TYPE "DT_ALM_SYSTEM_GEN_SPEED_WH_AND_VIB"
VERSION : 0.1
   STRUCT
      F1_ERR { S7_SetPoint := 'False'} : "DT_ALM_SOLO" := (192, FALSE, FALSE, TRUE, (), (), 2, 4, 2, (), (), (), (), (), T#3S);
      F1_H { S7_SetPoint := 'False'} : "DT_ALM_SOLO" := (193, FALSE, FALSE, TRUE, (), (), 2, 4, 1, (), (), (), (), (), T#5S);
      F1_HH { S7_SetPoint := 'False'} : "DT_ALM_SOLO" := (194, FALSE, FALSE, TRUE, (), (), 2, 4, 3, (), (), (), (), (), T#5S);
      F2_ERR { S7_SetPoint := 'False'} : "DT_ALM_SOLO" := (195, FALSE, FALSE, TRUE, (), (), 2, 4, 2, (), (), (), (), (), T#3S);
      F2_H { S7_SetPoint := 'False'} : "DT_ALM_SOLO" := (196, FALSE, FALSE, TRUE, (), (), 2, 4, 1, (), (), (), (), (), T#5S);
      F2_HH { S7_SetPoint := 'False'} : "DT_ALM_SOLO" := (197, FALSE, FALSE, TRUE, (), (), 2, 4, 3, (), (), (), (), (), T#5S);
      F3_ERR { S7_SetPoint := 'False'} : "DT_ALM_SOLO" := (198, FALSE, FALSE, FALSE, (), (), 0, 0, 0, (), (), (), (), (), T#500MS);
      F3_H { S7_SetPoint := 'False'} : "DT_ALM_SOLO" := (199, FALSE, FALSE, FALSE, (), (), 0, 0, 0, (), (), (), (), (), T#500MS);
      F3_HH { S7_SetPoint := 'False'} : "DT_ALM_SOLO" := (200, FALSE, FALSE, FALSE, (), (), 0, 0, 0, (), (), (), (), (), T#500MS);
      F4_ERR { S7_SetPoint := 'False'} : "DT_ALM_SOLO" := (201, FALSE, FALSE, TRUE, (), (), 2, 4, 2, (), (), (), (), (), T#3S);
      F4_H { S7_SetPoint := 'False'} : "DT_ALM_SOLO" := (202, FALSE, FALSE, TRUE, (), (), 2, 4, 1, (), (), (), (), (), T#5S);
      F4_HH { S7_SetPoint := 'False'} : "DT_ALM_SOLO" := (203, FALSE, FALSE, TRUE, (), (), 2, 4, 3, (), (), (), (), (), T#5S);
      SPARE_204 { S7_SetPoint := 'False'} : "DT_ALM_SOLO" := (204, FALSE, FALSE, FALSE, (), (), 0, 0, 0, (), (), (), (), (), T#500MS);
      SPARE_205 { S7_SetPoint := 'False'} : "DT_ALM_SOLO" := (205, FALSE, FALSE, FALSE, (), (), 0, 0, 0, (), (), (), (), (), T#500MS);
      SPARE_206 { S7_SetPoint := 'False'} : "DT_ALM_SOLO" := (206, FALSE, FALSE, FALSE, (), (), 0, 0, 0, (), (), (), (), (), T#500MS);
      SPARE_207 { S7_SetPoint := 'False'} : "DT_ALM_SOLO" := (207, FALSE, FALSE, FALSE, (), (), 0, 0, 0, (), (), (), (), (), T#500MS);
      WH_DE_1_W { S7_SetPoint := 'False'} : "DT_ALM_SOLO" := (208, FALSE, TRUE, TRUE, (), (), 0, 0, 1, (), (), (), (), (), T#500MS);
      WH_DE_1_T { S7_SetPoint := 'False'} : "DT_ALM_SOLO" := (209, FALSE, TRUE, TRUE, (), (), 0, 0, 2, (), (), (), (), (), T#500MS);
      WH_DE_2_W { S7_SetPoint := 'False'} : "DT_ALM_SOLO" := (210, FALSE, FALSE, FALSE, (), (), 0, 0, 0, (), (), (), (), (), T#500MS);
      WH_DE_2_T { S7_SetPoint := 'False'} : "DT_ALM_SOLO" := (211, FALSE, FALSE, FALSE, (), (), 0, 0, 0, (), (), (), (), (), T#500MS);
      WH_NDE_1_W { S7_SetPoint := 'False'} : "DT_ALM_SOLO" := (212, FALSE, TRUE, TRUE, (), (), 0, 0, 1, (), (), (), (), (), T#500MS);
      WH_NDE_1_T { S7_SetPoint := 'False'} : "DT_ALM_SOLO" := (213, FALSE, TRUE, TRUE, (), (), 0, 0, 2, (), (), (), (), (), T#500MS);
      WH_NDE_2_W { S7_SetPoint := 'False'} : "DT_ALM_SOLO" := (214, FALSE, FALSE, FALSE, (), (), 0, 0, 0, (), (), (), (), (), T#500MS);
      WH_NDE_2_T { S7_SetPoint := 'False'} : "DT_ALM_SOLO" := (215, FALSE, FALSE, FALSE, (), (), 0, 0, 0, (), (), (), (), (), T#500MS);
      SPEED_MAIN_ERR { S7_SetPoint := 'False'} : "DT_ALM_SOLO" := (216, FALSE, FALSE, FALSE, (), (), 0, 0, 0, (), (), (), (), (), T#500MS);
      SPEED_RED_ERR { S7_SetPoint := 'False'} : "DT_ALM_SOLO" := (217, FALSE, TRUE, TRUE, (), (), 2, 4, 2, (), (), (), (), (), T#3S);
      SPEED_DIFF_N1_N2 { S7_SetPoint := 'False'} : "DT_ALM_SOLO" := (218, FALSE, FALSE, FALSE, (), (), 0, 0, 0, (), (), (), (), (), T#500MS);
      SPEED_DIFF_N1_F { S7_SetPoint := 'False'} : "DT_ALM_SOLO" := (219, FALSE, TRUE, TRUE, (), (), 2, 0, 0, (), (), (), (), (), T#5S);
      SPEED_OVERSPEED1 { S7_SetPoint := 'False'} : "DT_ALM_SOLO" := (220, FALSE, TRUE, TRUE, (), (), 0, 0, 2, (), (), (), (), (), T#5S);
      SPEED_OVERSPEED2 { S7_SetPoint := 'False'} : "DT_ALM_SOLO" := (221, FALSE, TRUE, TRUE, (), (), 1, 0, 3, (), (), (), (), (), T#2S);
      SPARE_222 { S7_SetPoint := 'False'} : "DT_ALM_SOLO" := (222, FALSE, FALSE, FALSE, (), (), 0, 0, 0, (), (), (), (), (), T#500MS);
      SPARE_223 { S7_SetPoint := 'False'} : "DT_ALM_SOLO" := (223, FALSE, FALSE, FALSE, (), (), 0, 0, 0, (), (), (), (), (), T#500MS);
   END_STRUCT;

END_TYPE

